(* IEC 61131-3 sources: tsplc/examples/bottling-line/raw-st/src/capping, 2 files *)

(* ---- E_CapperState.st ---- *)
{attribute 'qualified_only'}
{attribute 'strict'}
TYPE E_CapperState : (Idle := 0, Capping := 1) USINT;
END_TYPE

(* ---- ST_Batch.st ---- *)
TYPE ST_Batch :
STRUCT
	Id : UDINT;
	CapTorques : ARRAY [1..4] OF REAL;
END_STRUCT
END_TYPE
